(* IEC 61131-3 sources: STruCpp/tests/st-validation/composite_access, 4 files *)

(* ---- nested_access.st ---- *)
TYPE Inner :
  STRUCT
    value : INT;
  END_STRUCT;
END_TYPE

TYPE Outer :
  STRUCT
    inner : Inner;
    count : INT;
  END_STRUCT;
END_TYPE

PROGRAM NestedAccessTest
  VAR
    data : Outer;
    result : INT;
  END_VAR

  data.inner.value := 42;
  data.count := 5;
  result := data.inner.value + data.count;
END_PROGRAM

(* ---- struct_member.st ---- *)
TYPE Point :
  STRUCT
    x : INT;
    y : INT;
  END_STRUCT;
END_TYPE

PROGRAM StructMemberTest
  VAR
    p : Point;
    dist : INT;
  END_VAR

  p.x := 3;
  p.y := 4;
  dist := p.x + p.y;
END_PROGRAM

(* ---- test_nested_access.st ---- *)
TEST 'Nested struct member access'
  VAR uut : NestedAccessTest; END_VAR
  uut();
  ASSERT_EQ(uut.data.inner.value, 42);
END_TEST

TEST 'Nested struct in expression'
  VAR uut : NestedAccessTest; END_VAR
  uut();
  ASSERT_EQ(uut.result, 47);
END_TEST

(* ---- test_struct_member.st ---- *)
TEST 'Struct member assignment'
  VAR uut : StructMemberTest; END_VAR
  uut();
  ASSERT_EQ(uut.p.x, 3);
  ASSERT_EQ(uut.p.y, 4);
END_TEST

TEST 'Struct member in expression'
  VAR uut : StructMemberTest; END_VAR
  uut();
  ASSERT_EQ(uut.dist, 7);
END_TEST
